Fanuc KAREL source: KT00626.KL

PROGRAM KT00626
%NOLOCKGROUP
VAR
  S1: STRING[80]
  S2: STRING[80]
  OUT: REAL
BEGIN
  S1 = 'A'
  S2 = 'B'
  S1 = 'A'
  S2 = 'B'
  OUT = NOT S1
END KT00626
